(* IEC 61131-3 sources: Antarbhukti-LLM/benchmarks, 12 files *)

(* ---- RISING_EDGE.st ---- *)
FUNCTION_BLOCK R_TRIG
VAR_INPUT CLK : BOOL; END_VAR
VAR_OUTPUT Q : BOOL; END_VAR
VAR state : INT := 0; END_VAR

CASE state OF
0: IF CLK THEN state := 1; END_IF;
1: Q := TRUE; state := 0;
END_CASE;
END_FUNCTION_BLOCK

(* ---- SR_LATCH.st ---- *)
FUNCTION_BLOCK SR
VAR_INPUT S : BOOL; R : BOOL; END_VAR
VAR_OUTPUT Q : BOOL; END_VAR
VAR state : INT := 0; END_VAR

CASE state OF
0: IF S THEN state := 1; END_IF;
1: IF R THEN state := 0; END_IF;
END_CASE;

Q := state = 1;
END_FUNCTION_BLOCK

(* ---- TOF.st ---- *)
FUNCTION_BLOCK TOF
VAR_INPUT
    IN : BOOL;
END_VAR
VAR_OUTPUT
    Q : BOOL;
END_VAR
VAR state : INT := 0; END_VAR

CASE state OF
0: IF NOT IN THEN state := 1; END_IF;
1: state := 2;
2: Q := FALSE;
END_CASE;
END_FUNCTION_BLOCK

(* ---- TON.st ---- *)
FUNCTION_BLOCK TON
VAR_INPUT
    IN : BOOL;
    PT : TIME;
END_VAR
VAR_OUTPUT
    Q : BOOL;
END_VAR
VAR
    state : INT := 0;
END_VAR

CASE state OF
0: IF IN THEN state := 1; END_IF;
1: state := 2;
2: Q := TRUE;
END_CASE;
END_FUNCTION_BLOCK

(* ---- BATCH_REACTOR.st ---- *)
PROGRAM REACTOR
VAR state : INT := 0; start : BOOL; END_VAR

CASE state OF
0: IF start THEN state := 1; END_IF;
1: state := 2;
2: state := 3;
3: state := 4;
4: state := 5;
5: state := 0;
END_CASE;
END_PROGRAM

(* ---- CONVEYOR_EMERGENCY.st ---- *)
PROGRAM CONVEYOR
VAR state : INT := 0; start : BOOL; emergency : BOOL; END_VAR

CASE state OF
0: IF start THEN state := 1; END_IF;
1: IF emergency THEN state := 3 ELSE state := 2; END_IF;
2: IF emergency THEN state := 3; END_IF;
3: state := 0;
END_CASE;
END_PROGRAM

(* ---- ELEVATOR_2FLOOR.st ---- *)
PROGRAM ELEVATOR
VAR state : INT := 0; call_up : BOOL; call_down : BOOL; END_VAR

CASE state OF
0: IF call_up THEN state := 1; END_IF;
1: state := 2;
2: state := 3;
3: IF call_down THEN state := 4; END_IF;
4: state := 0;
END_CASE;
END_PROGRAM

(* ---- MODE_MANAGER.st ---- *)
PROGRAM MODE_MANAGER
VAR state : INT := 0; auto : BOOL; fault : BOOL; END_VAR

CASE state OF
0: IF auto THEN state := 1; END_IF;
1: IF fault THEN state := 3; END_IF;
3: state := 2;
2: state := 0;
END_CASE;
END_PROGRAM

(* ---- PICK_PLACE_ROBOT.st ---- *)
PROGRAM PICK_PLACE
VAR state : INT := 0; part_ready : BOOL; END_VAR

CASE state OF
0: IF part_ready THEN state := 1; END_IF;
1: state := 2;
2: state := 3;
3: state := 4;
4: state := 5;
5: state := 0;
END_CASE;
END_PROGRAM

(* ---- TANK_FILLING.st ---- *)
PROGRAM TANK
VAR state : INT := 0; low : BOOL; high : BOOL; END_VAR

CASE state OF
0: IF low THEN state := 1; END_IF;
1: IF high THEN state := 2; END_IF;
2: state := 3;
3: state := 0;
END_CASE;
END_PROGRAM

(* ---- TRAFFIC_LIGHT.st ---- *)
PROGRAM TRAFFIC_LIGHT
VAR state : INT := 0; END_VAR

CASE state OF
0: state := 1;
1: state := 2;
2: state := 3;
3: state := 0;
END_CASE;
END_PROGRAM

(* ---- WASHING_MACHINE.st ---- *)
PROGRAM WASHING_MACHINE
VAR state : INT := 0; start : BOOL; END_VAR

CASE state OF
0: IF start THEN state := 1; END_IF;
1: state := 2;
2: state := 3;
3: state := 4;
4: state := 5;
5: state := 0;
END_CASE;
END_PROGRAM
